(*
SPDX-FileCopyrightText: © 2026 Oleksandr Tiutyk <trofimich@gmail.com>
SPDX-License-Identifier: MIT
License: https://opensource.org/license/mit
*)

(*!
<summary>Reports the outcome of a single running step in Activity.OnRunning.</summary>
<description>
WORK_IN_PROGRESS keeps the activity in ACTIVE_RUNNING for subsequent Execute calls. WORK_COMPLETED transitions
the activity to PASSIVE_COMPLETED. WORK_HALTED transitions the activity to PASSIVE_HALTED and requires a
non-whitespace haltReason output.
</description>
*)

{attribute 'qualified_only'}
{attribute 'strict'}
{attribute 'to_string'}
TYPE ACTIVITY_RUNNING_STATE :
(
	WORK_IN_PROGRESS := 0,
	WORK_COMPLETED,
	WORK_HALTED
);
END_TYPE

(* stored: Version 1.1.0.1
   DUT ACTIVITY_RUNNING_STATE: Id {24d4d980-d91a-4e70-b1c0-2be206ebd59f} *)
